// TwinCAT 3 PLC project TestRunner
// Title: TestRunner
// Company: Intecre Ltd
// ProjectVersion: 1.0.0.0
// Description: TcUnit test suites for the Intecre.File library. Not a library; activate it on a runtime (the usermode runtime works) to run the tests. The tests write their files to C:\TcUnit_IntecreFile.
// ProgramVersion: 3.1.4026.25
// libraries:
//   Tc2_Standard, * (Beckhoff Automation GmbH)
//   Tc2_System, * (Beckhoff Automation GmbH)
//   Tc2_Utilities, * (Beckhoff Automation GmbH)
//   TcUnit, * (www.tcunit.org)
//   Intecre.File, * (Intecre Ltd)
// project tree:
//   / MAIN.TcPOU, PlcTask.TcTTO
//   Helpers/ F_TestFilePath.TcPOU, ST_TestRecipe.TcDUT, T_TestDirectory.TcPOU, T_TestFile.TcPOU, TestFiles.TcGVL
//   Tests/ T_TxtFileWriter_Tests.TcPOU, T_CsvFileWriter_Tests.TcPOU, T_CsvFileReader_Tests.TcPOU, T_StructJsonFile_Tests.TcPOU, T_StructPersistence_Tests.TcPOU, T_CheckFileExists_Tests.TcPOU, ProjectInformation_Tests.TcPOU
// (motion and I/O tree: see PLC project intecre_file)
// real-time tasks:
//   TASK PlcTask: cycle T#10ms, priority 20, ADS port 350

CONFIGURATION TestRunner
    RESOURCE PLC ON TwinCAT3
        TASK PlcTask(INTERVAL := T#10ms, PRIORITY := 20);
        PROGRAM MAIN WITH PlcTask : MAIN;
    END_RESOURCE
END_CONFIGURATION

// ---- Helpers/ST_TestRecipe.TcDUT
TYPE ST_TestRecipe :
STRUCT
  Name : STRING(40);
  Speed : LREAL;
  Count : DINT;
  Enabled : BOOL;
END_STRUCT
END_TYPE

// ---- Helpers/TestFiles.TcGVL
{attribute 'qualified_only'}
VAR_GLOBAL CONSTANT
  DIRECTORY : T_MaxString := 'C:\TcUnit_IntecreFile';
  TIMEOUT : TIME := T#5S;
END_VAR

// ---- MAIN.TcPOU
PROGRAM MAIN
VAR
  testDirectory           : T_TestDirectory;
  suiteTxtFileWriter      : T_TxtFileWriter_Tests;
  suiteCsvFileWriter      : T_CsvFileWriter_Tests;
  suiteCsvFileReader      : T_CsvFileReader_Tests;
  suiteStructJsonFile     : T_StructJsonFile_Tests;
  suiteStructPersistence  : T_StructPersistence_Tests;
  suiteCheckFileExists    : T_CheckFileExists_Tests;
  suiteProjectInformation : ProjectInformation_Tests;
END_VAR

testDirectory();

IF NOT testDirectory.Ready THEN
  RETURN;
END_IF

TcUnit.RUN_IN_SEQUENCE();

END_PROGRAM

// ---- Helpers/T_TestDirectory.TcPOU
FUNCTION_BLOCK T_TestDirectory
VAR
  createDirectory : FB_CreateDir;
  requested : BOOL;
  _ready : BOOL;
END_VAR

IF _ready THEN
  RETURN;
END_IF

createDirectory(sNetId := '', sPathName := TestFiles.DIRECTORY, bExecute := TRUE);

IF requested AND NOT createDirectory.bBusy THEN
  _ready := TRUE;
END_IF

requested := TRUE;

PROPERTY Ready : BOOL
GET
Ready := _ready;
END_GET
END_PROPERTY

END_FUNCTION_BLOCK

// ---- Tests/T_TxtFileWriter_Tests.TcPOU
FUNCTION_BLOCK T_TxtFileWriter_Tests EXTENDS TcUnit.FB_TestSuite

Test_WriteLineEndsEachLineWithCrlf();
Test_WriteAddsToTheCurrentLine();
Test_AppendModeAddsToTheEndOfTheFile();
Test_OverwriteModeReplacesTheFile();
Test_ClearBufferDiscardsWhatWasWritten();
Test_ClearBufferReportsTheBufferIsClear();
Test_KeepsLinesLongerThan255Characters();
Test_MissingDirectoryGivesAnError();

METHOD PRIVATE Test_WriteLineEndsEachLineWithCrlf
VAR_INST
  writer : T_TxtFileWriter;
  testFile : T_TestFile;
  timeout : TON;
  step : INT;
END_VAR
IF NOT TcUnit.TEST_ORDERED(__POUNAME()) THEN
  RETURN;
END_IF

writer();
testFile();

timeout(IN := TRUE, PT := TestFiles.TIMEOUT);

IF timeout.Q THEN
  AssertTrue(Condition := FALSE, Message := 'the file operation did not finish in time');
  TEST_FINISHED_NAMED(__POUNAME());
  RETURN;
END_IF

CASE step OF

  0:

    writer.SetFileParams(FilePath := F_TestFilePath('txt_write_line.txt'));
    writer.WriteLine(Entry := 'first');
    writer.WriteLine(Entry := 'second');
    writer.WriteToFile();
    step := 10;

  10:

    IF writer.Busy THEN
      RETURN;
    END_IF

    AssertFalse(Condition := writer.Error, Message := 'file written without an error');
    testFile.Read(FilePath := F_TestFilePath('txt_write_line.txt'));
    step := 20;

  20:

    IF testFile.Busy THEN
      RETURN;
    END_IF

    AssertEquals_STRING(Expected := 'first$R$Nsecond$R$N', Actual := testFile.Text, Message := 'each line ends with CR LF');
    TEST_FINISHED_NAMED(__POUNAME());

END_CASE
END_METHOD

METHOD PRIVATE Test_WriteAddsToTheCurrentLine
VAR_INST
  writer : T_TxtFileWriter;
  testFile : T_TestFile;
  timeout : TON;
  step : INT;
END_VAR
IF NOT TcUnit.TEST_ORDERED(__POUNAME()) THEN
  RETURN;
END_IF

writer();
testFile();

timeout(IN := TRUE, PT := TestFiles.TIMEOUT);

IF timeout.Q THEN
  AssertTrue(Condition := FALSE, Message := 'the file operation did not finish in time');
  TEST_FINISHED_NAMED(__POUNAME());
  RETURN;
END_IF

CASE step OF

  0:

    writer.SetFileParams(FilePath := F_TestFilePath('txt_write.txt'));
    writer.Write(Entry := 'one');
    writer.Write(Entry := 'two');
    writer.NewLine();
    writer.WriteToFile();
    step := 10;

  10:

    IF writer.Busy THEN
      RETURN;
    END_IF

    AssertFalse(Condition := writer.Error, Message := 'file written without an error');
    testFile.Read(FilePath := F_TestFilePath('txt_write.txt'));
    step := 20;

  20:

    IF testFile.Busy THEN
      RETURN;
    END_IF

    AssertEquals_STRING(Expected := 'onetwo$R$N', Actual := testFile.Text, Message := 'Write adds to the line, NewLine ends it');
    TEST_FINISHED_NAMED(__POUNAME());

END_CASE
END_METHOD

METHOD PRIVATE Test_AppendModeAddsToTheEndOfTheFile
VAR_INST
  writer : T_TxtFileWriter;
  testFile : T_TestFile;
  timeout : TON;
  step : INT;
END_VAR
IF NOT TcUnit.TEST_ORDERED(__POUNAME()) THEN
  RETURN;
END_IF

writer();
testFile();

timeout(IN := TRUE, PT := TestFiles.TIMEOUT);

IF timeout.Q THEN
  AssertTrue(Condition := FALSE, Message := 'the file operation did not finish in time');
  TEST_FINISHED_NAMED(__POUNAME());
  RETURN;
END_IF

CASE step OF

  0:

    testFile.Write(FilePath := F_TestFilePath('txt_append.txt'), Content := 'existing$R$N');
    step := 5;

  5:

    IF testFile.Busy THEN
      RETURN;
    END_IF

    AssertFalse(Condition := testFile.Error, Message := 'existing file written');
    step := 6;

  6:

    writer.SetFileParams(FilePath := F_TestFilePath('txt_append.txt'));
    writer.SetFileOpenMode(Append := TRUE);
    writer.WriteLine(Entry := 'added');
    writer.WriteToFile();
    step := 10;

  10:

    IF writer.Busy THEN
      RETURN;
    END_IF

    AssertFalse(Condition := writer.Error, Message := 'file written without an error');
    testFile.Read(FilePath := F_TestFilePath('txt_append.txt'));
    step := 20;

  20:

    IF testFile.Busy THEN
      RETURN;
    END_IF

    AssertEquals_STRING(Expected := 'existing$R$Nadded$R$N', Actual := testFile.Text, Message := 'appended after the existing line');
    TEST_FINISHED_NAMED(__POUNAME());

END_CASE
END_METHOD

METHOD PRIVATE Test_OverwriteModeReplacesTheFile
VAR_INST
  writer : T_TxtFileWriter;
  testFile : T_TestFile;
  timeout : TON;
  step : INT;
END_VAR
IF NOT TcUnit.TEST_ORDERED(__POUNAME()) THEN
  RETURN;
END_IF

writer();
testFile();

timeout(IN := TRUE, PT := TestFiles.TIMEOUT);

IF timeout.Q THEN
  AssertTrue(Condition := FALSE, Message := 'the file operation did not finish in time');
  TEST_FINISHED_NAMED(__POUNAME());
  RETURN;
END_IF

CASE step OF

  0:

    testFile.Write(FilePath := F_TestFilePath('txt_overwrite.txt'), Content := 'old content$R$N');
    step := 5;

  5:

    IF testFile.Busy THEN
      RETURN;
    END_IF

    AssertFalse(Condition := testFile.Error, Message := 'existing file written');
    step := 6;

  6:

    writer.SetFileParams(FilePath := F_TestFilePath('txt_overwrite.txt'));
    writer.WriteLine(Entry := 'new');
    writer.WriteToFile();
    step := 10;

  10:

    IF writer.Busy THEN
      RETURN;
    END_IF

    AssertFalse(Condition := writer.Error, Message := 'file written without an error');
    testFile.Read(FilePath := F_TestFilePath('txt_overwrite.txt'));
    step := 20;

  20:

    IF testFile.Busy THEN
      RETURN;
    END_IF

    AssertEquals_STRING(Expected := 'new$R$N', Actual := testFile.Text, Message := 'the old content is gone');
    TEST_FINISHED_NAMED(__POUNAME());

END_CASE
END_METHOD

METHOD PRIVATE Test_ClearBufferDiscardsWhatWasWritten
VAR_INST
  writer : T_TxtFileWriter;
  testFile : T_TestFile;
  timeout : TON;
  step : INT;
END_VAR
IF NOT TcUnit.TEST_ORDERED(__POUNAME()) THEN
  RETURN;
END_IF

writer();
testFile();

timeout(IN := TRUE, PT := TestFiles.TIMEOUT);

IF timeout.Q THEN
  AssertTrue(Condition := FALSE, Message := 'the file operation did not finish in time');
  TEST_FINISHED_NAMED(__POUNAME());
  RETURN;
END_IF

CASE step OF

  0:

    writer.SetFileParams(FilePath := F_TestFilePath('txt_clear_buffer.txt'));
    writer.WriteLine(Entry := 'discarded');
    writer.ClearBuffer();
    writer.WriteLine(Entry := 'kept');
    writer.WriteToFile();
    step := 10;

  10:

    IF writer.Busy THEN
      RETURN;
    END_IF

    AssertFalse(Condition := writer.Error, Message := 'file written without an error');
    testFile.Read(FilePath := F_TestFilePath('txt_clear_buffer.txt'));
    step := 20;

  20:

    IF testFile.Busy THEN
      RETURN;
    END_IF

    AssertEquals_STRING(Expected := 'kept$R$N', Actual := testFile.Text, Message := 'only the line written after ClearBuffer');
    TEST_FINISHED_NAMED(__POUNAME());

END_CASE
END_METHOD

METHOD PRIVATE Test_ClearBufferReportsTheBufferIsClear
VAR_INST
  writer : T_TxtFileWriter;
END_VAR
IF NOT TcUnit.TEST_ORDERED(__POUNAME()) THEN
  RETURN;
END_IF

writer.WriteLine(Entry := 'line');
AssertTrue(Condition := writer.ClearBuffer(), Message := 'ClearBuffer returns TRUE');
AssertTrue(Condition := writer.BufferClear, Message := 'BufferClear after ClearBuffer');

TEST_FINISHED_NAMED(__POUNAME());
END_METHOD

METHOD PRIVATE Test_KeepsLinesLongerThan255Characters
VAR_INST
  writer : T_TxtFileWriter;
  testFile : T_TestFile;
  timeout : TON;
  step : INT;
  longLine : TxtFileString;
END_VAR
IF NOT TcUnit.TEST_ORDERED(__POUNAME()) THEN
  RETURN;
END_IF

writer();
testFile();

timeout(IN := TRUE, PT := TestFiles.TIMEOUT);

IF timeout.Q THEN
  AssertTrue(Condition := FALSE, Message := 'the file operation did not finish in time');
  TEST_FINISHED_NAMED(__POUNAME());
  RETURN;
END_IF

CASE step OF

  0:

    MEMSET(destAddr := ADR(longLine), fillByte := 16#41, n := 300);
    writer.SetFileParams(FilePath := F_TestFilePath('txt_long_line.txt'));
    writer.WriteLine(Entry := longLine);
    writer.WriteToFile();
    step := 10;

  10:

    IF writer.Busy THEN
      RETURN;
    END_IF

    testFile.Read(FilePath := F_TestFilePath('txt_long_line.txt'));
    step := 20;

  20:

    IF testFile.Busy THEN
      RETURN;
    END_IF

    AssertEquals_DINT(Expected := 302, Actual := testFile.Length, Message := '300 characters and CR LF');
    TEST_FINISHED_NAMED(__POUNAME());

END_CASE
END_METHOD

METHOD PRIVATE Test_MissingDirectoryGivesAnError
VAR_INST
  writer : T_TxtFileWriter;
  timeout : TON;
  step : INT;
END_VAR
IF NOT TcUnit.TEST_ORDERED(__POUNAME()) THEN
  RETURN;
END_IF

writer();

timeout(IN := TRUE, PT := TestFiles.TIMEOUT);

IF timeout.Q THEN
  AssertTrue(Condition := FALSE, Message := 'the file operation did not finish in time');
  TEST_FINISHED_NAMED(__POUNAME());
  RETURN;
END_IF

CASE step OF

  0:

    writer.SetFileParams(FilePath := F_TestFilePath('missing\file.txt'));
    writer.WriteLine(Entry := 'line');
    writer.WriteToFile();
    step := 10;

  10:

    IF writer.Busy THEN
      RETURN;
    END_IF

    AssertTrue(Condition := writer.Error, Message := 'a folder that does not exist gives an error');
    AssertTrue(Condition := writer.ErrorId <> 0, Message := 'with an error id');
    TEST_FINISHED_NAMED(__POUNAME());

END_CASE
END_METHOD

END_FUNCTION_BLOCK

// ---- Helpers/T_TestFile.TcPOU
FUNCTION_BLOCK T_TestFile
VAR
  fileOpen : FB_FileOpen;
  fileWrite : FB_FileWrite;
  fileRead : FB_FileRead;
  fileClose : FB_FileClose;
  fileDelete : FB_FileDelete;
  path : T_MaxString;
  textToWrite : STRING(2000);
  textRead : STRING(2000);
  startOfTextRead : T_MaxString;
  bytesRead : UDINT;
  request : (NoRequest, WriteRequest, ReadRequest, DeleteRequest);
  state : (Idle, Opening, Writing, Reading, Closing, Deleting);
  failed : BOOL;
END_VAR

CASE state OF

  Idle:

    IF request = DeleteRequest THEN
      state := Deleting;

    ELSIF request <> NoRequest THEN
      state := Opening;

    END_IF

  Opening:

    IF NOT fileOpen.bBusy AND fileOpen.bError THEN
      Finish(WithError := TRUE);

    ELSIF NOT fileOpen.bBusy AND (request = WriteRequest) THEN
      state := Writing;

    ELSIF NOT fileOpen.bBusy THEN
      state := Reading;

    END_IF

  Writing:

    IF NOT fileWrite.bBusy THEN
      failed := fileWrite.bError;
      state := Closing;
    END_IF

  Reading:

    IF NOT fileRead.bBusy THEN
      failed := fileRead.bError;
      bytesRead := fileRead.cbRead;
      MEMCPY(destAddr := ADR(startOfTextRead), srcAddr := ADR(textRead), n := SIZEOF(startOfTextRead) - 1);
      state := Closing;
    END_IF

  Closing:

    IF NOT fileClose.bBusy THEN
      Finish(WithError := failed OR fileClose.bError);
    END_IF

  Deleting:

    IF NOT fileDelete.bBusy THEN
      Finish(WithError := fileDelete.bError);
    END_IF

END_CASE

fileOpen(
  sNetId := '',
  sPathName := path,
  nMode := SEL(request = WriteRequest, FOPEN_MODEREAD OR FOPEN_MODEBINARY, FOPEN_MODEWRITE OR FOPEN_MODEBINARY),
  bExecute := state = Opening);

fileWrite(
  sNetId := '',
  hFile := fileOpen.hFile,
  pWriteBuff := ADR(textToWrite),
  cbWriteLen := TO_UDINT(LEN2(ADR(textToWrite))),
  bExecute := state = Writing);

fileRead(
  sNetId := '',
  hFile := fileOpen.hFile,
  pReadBuff := ADR(textRead),
  cbReadLen := SIZEOF(textRead) - 1,
  bExecute := state = Reading);

fileClose(
  sNetId := '',
  hFile := fileOpen.hFile,
  bExecute := state = Closing);

fileDelete(
  sNetId := '',
  sPathName := path,
  bExecute := state = Deleting);

PROPERTY Busy : BOOL
GET
Busy := request <> NoRequest;
END_GET
END_PROPERTY

METHOD Contains : BOOL
VAR_INPUT
  Part : T_MaxString;
END_VAR
VAR
  textLength : DINT;
  partLength : DINT;
  position : DINT;
END_VAR
textLength := TO_DINT(LEN2(ADR(textRead)));
partLength := TO_DINT(LEN2(ADR(Part)));

IF partLength = 0 THEN
  RETURN;
END_IF

FOR position := 0 TO textLength - partLength DO
  IF MEMCMP(pBuf1 := ADR(textRead) + TO_UDINT(position), pBuf2 := ADR(Part), n := TO_UDINT(partLength)) = 0 THEN
    Contains := TRUE;
    RETURN;
  END_IF
END_FOR
END_METHOD

METHOD Delete : BOOL
VAR_INPUT
  FilePath : T_MaxString;
END_VAR
IF Busy THEN
  RETURN;
END_IF

path := FilePath;
failed := FALSE;
request := DeleteRequest;
Delete := TRUE;
END_METHOD

PROPERTY Error : BOOL
GET
Error := failed AND NOT Busy;
END_GET
END_PROPERTY

METHOD PRIVATE Finish
VAR_INPUT
  WithError : BOOL;
END_VAR
failed := WithError;
request := NoRequest;
state := Idle;
END_METHOD

PROPERTY LastByte : BYTE // the last byte of the file the last Read read; 0 when it read nothing
GET // PUBLIC
IF bytesRead = 0 THEN
  RETURN;
END_IF

LastByte := textRead[bytesRead - 1];
END_GET
END_PROPERTY

PROPERTY Length : DINT
GET
Length := TO_DINT(LEN2(ADR(textRead)));
END_GET
END_PROPERTY

METHOD Read : BOOL
VAR_INPUT
  FilePath : T_MaxString;
END_VAR
IF Busy THEN
  RETURN;
END_IF

path := FilePath;
MEMSET(destAddr := ADR(textRead), fillByte := 0, n := SIZEOF(textRead));
MEMSET(destAddr := ADR(startOfTextRead), fillByte := 0, n := SIZEOF(startOfTextRead));
bytesRead := 0;
failed := FALSE;
request := ReadRequest;
Read := TRUE;
END_METHOD

PROPERTY Text : T_MaxString
GET
Text := startOfTextRead;
END_GET
END_PROPERTY

METHOD Write : BOOL
VAR_INPUT
  FilePath : T_MaxString;
  Content : STRING(2000);
END_VAR
IF Busy THEN
  RETURN;
END_IF

path := FilePath;
textToWrite := Content;
failed := FALSE;
request := WriteRequest;
Write := TRUE;
END_METHOD

END_FUNCTION_BLOCK

// ---- Helpers/F_TestFilePath.TcPOU
FUNCTION F_TestFilePath : T_MaxString
VAR_INPUT
  FileName : T_MaxString;
END_VAR

F_TestFilePath := CONCAT(CONCAT(TestFiles.DIRECTORY, '\'), FileName);

END_FUNCTION

// ---- Tests/T_CsvFileWriter_Tests.TcPOU
FUNCTION_BLOCK T_CsvFileWriter_Tests EXTENDS TcUnit.FB_TestSuite

Test_SeparatesFieldsWithCommas();
Test_SeparatesFieldsWithSemicolons();
Test_UnknownSeparatorFallsBackToSemicolon();
Test_AppendModeAddsRows();
Test_QuotesAFieldContainingTheSeparator();
Test_CountsRowsAndColumns();
Test_ClearBufferReportsTheBufferIsClear();

METHOD PRIVATE Test_SeparatesFieldsWithCommas
VAR_INST
  writer : T_CsvFileWriter;
  testFile : T_TestFile;
  timeout : TON;
  step : INT;
END_VAR
IF NOT TcUnit.TEST_ORDERED(__POUNAME()) THEN
  RETURN;
END_IF

writer();
testFile();

timeout(IN := TRUE, PT := TestFiles.TIMEOUT);

IF timeout.Q THEN
  AssertTrue(Condition := FALSE, Message := 'the file operation did not finish in time');
  TEST_FINISHED_NAMED(__POUNAME());
  RETURN;
END_IF

CASE step OF

  0:

    writer.SetFileParams(FilePath := F_TestFilePath('csv_commas.csv'), Separator := ASCI_COMMA);
    writer.AddStringField(sFieldString := 'a');
    writer.AddStringField(sFieldString := 'b');
    writer.NewLine();
    writer.AddStringField(sFieldString := 'c');
    writer.AddStringField(sFieldString := 'd');
    writer.WriteToFile();
    step := 10;

  10:

    IF writer.Busy THEN
      RETURN;
    END_IF

    AssertFalse(Condition := writer.Error, Message := 'file written without an error');
    testFile.Read(FilePath := F_TestFilePath('csv_commas.csv'));
    step := 20;

  20:

    IF testFile.Busy THEN
      RETURN;
    END_IF

    AssertEquals_STRING(Expected := 'a,b$R$Nc,d$R$N', Actual := testFile.Text, Message := 'two rows of two comma separated fields');
    TEST_FINISHED_NAMED(__POUNAME());

END_CASE
END_METHOD

METHOD PRIVATE Test_SeparatesFieldsWithSemicolons
VAR_INST
  writer : T_CsvFileWriter;
  testFile : T_TestFile;
  timeout : TON;
  step : INT;
END_VAR
IF NOT TcUnit.TEST_ORDERED(__POUNAME()) THEN
  RETURN;
END_IF

writer();
testFile();

timeout(IN := TRUE, PT := TestFiles.TIMEOUT);

IF timeout.Q THEN
  AssertTrue(Condition := FALSE, Message := 'the file operation did not finish in time');
  TEST_FINISHED_NAMED(__POUNAME());
  RETURN;
END_IF

CASE step OF

  0:

    writer.SetFileParams(FilePath := F_TestFilePath('csv_semicolons.csv'), Separator := ASCI_SEMI_COLON);
    writer.AddStringField(sFieldString := 'a');
    writer.AddStringField(sFieldString := 'b');
    writer.WriteToFile();
    step := 10;

  10:

    IF writer.Busy THEN
      RETURN;
    END_IF

    AssertFalse(Condition := writer.Error, Message := 'file written without an error');
    testFile.Read(FilePath := F_TestFilePath('csv_semicolons.csv'));
    step := 20;

  20:

    IF testFile.Busy THEN
      RETURN;
    END_IF

    AssertEquals_STRING(Expected := 'a;b$R$N', Actual := testFile.Text, Message := 'semicolon separated fields');
    TEST_FINISHED_NAMED(__POUNAME());

END_CASE
END_METHOD

METHOD PRIVATE Test_UnknownSeparatorFallsBackToSemicolon
VAR_INST
  writer : T_CsvFileWriter;
  testFile : T_TestFile;
  timeout : TON;
  step : INT;
END_VAR
IF NOT TcUnit.TEST_ORDERED(__POUNAME()) THEN
  RETURN;
END_IF

writer();
testFile();

timeout(IN := TRUE, PT := TestFiles.TIMEOUT);

IF timeout.Q THEN
  AssertTrue(Condition := FALSE, Message := 'the file operation did not finish in time');
  TEST_FINISHED_NAMED(__POUNAME());
  RETURN;
END_IF

CASE step OF

  0:

    writer.SetFileParams(FilePath := F_TestFilePath('csv_unknown_separator.csv'), Separator := 16#09);
    writer.AddStringField(sFieldString := 'a');
    writer.AddStringField(sFieldString := 'b');
    writer.WriteToFile();
    step := 10;

  10:

    IF writer.Busy THEN
      RETURN;
    END_IF

    AssertFalse(Condition := writer.Error, Message := 'file written without an error');
    testFile.Read(FilePath := F_TestFilePath('csv_unknown_separator.csv'));
    step := 20;

  20:

    IF testFile.Busy THEN
      RETURN;
    END_IF

    AssertEquals_STRING(Expected := 'a;b$R$N', Actual := testFile.Text, Message := 'a tab is not supported, so semicolon is used');
    TEST_FINISHED_NAMED(__POUNAME());

END_CASE
END_METHOD

METHOD PRIVATE Test_AppendModeAddsRows
VAR_INST
  writer : T_CsvFileWriter;
  testFile : T_TestFile;
  timeout : TON;
  step : INT;
END_VAR
IF NOT TcUnit.TEST_ORDERED(__POUNAME()) THEN
  RETURN;
END_IF

writer();
testFile();

timeout(IN := TRUE, PT := TestFiles.TIMEOUT);

IF timeout.Q THEN
  AssertTrue(Condition := FALSE, Message := 'the file operation did not finish in time');
  TEST_FINISHED_NAMED(__POUNAME());
  RETURN;
END_IF

CASE step OF

  0:

    testFile.Write(FilePath := F_TestFilePath('csv_append.csv'), Content := 'x,y$R$N');
    step := 5;

  5:

    IF testFile.Busy THEN
      RETURN;
    END_IF

    AssertFalse(Condition := testFile.Error, Message := 'existing file written');
    step := 6;

  6:

    writer.SetFileParams(FilePath := F_TestFilePath('csv_append.csv'), Separator := ASCI_COMMA);
    writer.SetFileOpenMode(Append := TRUE);
    writer.AddStringField(sFieldString := 'a');
    writer.AddStringField(sFieldString := 'b');
    writer.WriteToFile();
    step := 10;

  10:

    IF writer.Busy THEN
      RETURN;
    END_IF

    AssertFalse(Condition := writer.Error, Message := 'file written without an error');
    testFile.Read(FilePath := F_TestFilePath('csv_append.csv'));
    step := 20;

  20:

    IF testFile.Busy THEN
      RETURN;
    END_IF

    AssertEquals_STRING(Expected := 'x,y$R$Na,b$R$N', Actual := testFile.Text, Message := 'row appended after the existing row');
    TEST_FINISHED_NAMED(__POUNAME());

END_CASE
END_METHOD

METHOD PRIVATE Test_QuotesAFieldContainingTheSeparator
VAR_INST
  writer : T_CsvFileWriter;
  testFile : T_TestFile;
  timeout : TON;
  step : INT;
END_VAR
IF NOT TcUnit.TEST_ORDERED(__POUNAME()) THEN
  RETURN;
END_IF

writer();
testFile();

timeout(IN := TRUE, PT := TestFiles.TIMEOUT);

IF timeout.Q THEN
  AssertTrue(Condition := FALSE, Message := 'the file operation did not finish in time');
  TEST_FINISHED_NAMED(__POUNAME());
  RETURN;
END_IF

CASE step OF

  0:

    writer.SetFileParams(FilePath := F_TestFilePath('csv_quoted.csv'), Separator := ASCI_COMMA);
    writer.AddStringField(sFieldString := 'a,b');
    writer.AddStringField(sFieldString := 'c');
    writer.WriteToFile();
    step := 10;

  10:

    IF writer.Busy THEN
      RETURN;
    END_IF

    AssertFalse(Condition := writer.Error, Message := 'file written without an error');
    testFile.Read(FilePath := F_TestFilePath('csv_quoted.csv'));
    step := 20;

  20:

    IF testFile.Busy THEN
      RETURN;
    END_IF

    AssertEquals_STRING(Expected := '"a,b",c$R$N', Actual := testFile.Text, Message := 'a field holding the separator is quoted so the row keeps two fields');
    TEST_FINISHED_NAMED(__POUNAME());

END_CASE
END_METHOD

METHOD PRIVATE Test_CountsRowsAndColumns
VAR_INST
  writer : T_CsvFileWriter;
END_VAR
IF NOT TcUnit.TEST_ORDERED(__POUNAME()) THEN
  RETURN;
END_IF

writer.SetFileParams(FilePath := F_TestFilePath('csv_counts.csv'), Separator := ASCI_COMMA);
writer.AddStringField(sFieldString := 'a');
writer.AddStringField(sFieldString := 'b');
AssertEquals_UINT(Expected := 2, Actual := writer.Column, Message := 'two fields on the row');
AssertEquals_UINT(Expected := 0, Actual := writer.Row, Message := 'still on the first row');

writer.NewLine();
AssertEquals_UINT(Expected := 0, Actual := writer.Column, Message := 'column back to zero on a new line');
AssertEquals_UINT(Expected := 1, Actual := writer.Row, Message := 'second row');

TEST_FINISHED_NAMED(__POUNAME());
END_METHOD

METHOD PRIVATE Test_ClearBufferReportsTheBufferIsClear
VAR_INST
  writer : T_CsvFileWriter;
END_VAR
IF NOT TcUnit.TEST_ORDERED(__POUNAME()) THEN
  RETURN;
END_IF

writer.SetFileParams(FilePath := F_TestFilePath('csv_clear.csv'), Separator := ASCI_COMMA);
writer.AddStringField(sFieldString := 'a');
AssertTrue(Condition := writer.ClearBuffer(), Message := 'ClearBuffer returns TRUE');
AssertTrue(Condition := writer.BufferClear, Message := 'BufferClear after ClearBuffer');

TEST_FINISHED_NAMED(__POUNAME());
END_METHOD

END_FUNCTION_BLOCK

// ---- Tests/T_CsvFileReader_Tests.TcPOU
FUNCTION_BLOCK T_CsvFileReader_Tests EXTENDS TcUnit.FB_TestSuite

Test_ReadsEachFieldWithItsRowAndColumn();
Test_ReadsSemicolonSeparatedFields();
Test_KeepsFieldsLongerThan80Characters();
Test_MissingFileGivesAnError();

METHOD PRIVATE Test_KeepsFieldsLongerThan80Characters
VAR_INST
  reader : T_CsvFileReader;
  testFile : T_TestFile;
  timeout : TON;
  step : INT;
  content : STRING(2000);
  field : T_MaxString;
END_VAR
IF NOT TcUnit.TEST_ORDERED(__POUNAME()) THEN
  RETURN;
END_IF

reader();
testFile();

timeout(IN := TRUE, PT := TestFiles.TIMEOUT);

IF timeout.Q THEN
  AssertTrue(Condition := FALSE, Message := 'the file operation did not finish in time');
  TEST_FINISHED_NAMED(__POUNAME());
  RETURN;
END_IF

CASE step OF

  0:

    MEMSET(destAddr := ADR(content), fillByte := 16#41, n := 100);
    content[100] := 16#0D;
    content[101] := 16#0A;
    testFile.Write(FilePath := F_TestFilePath('csv_long_field.csv'), Content := content);
    step := 10;

  10:

    IF testFile.Busy THEN
      RETURN;
    END_IF

    AssertFalse(Condition := testFile.Error, Message := 'CSV file written for the test');
    reader.SetFileParams(FilePath := F_TestFilePath('csv_long_field.csv'), Separator := ASCI_COMMA);
    reader.GetFile();
    step := 20;

  20:

    IF reader.Busy THEN
      RETURN;
    END_IF

    AssertFalse(Condition := reader.Error, Message := 'file read without an error');
    AssertTrue(Condition := reader.ReadyForParsing, Message := 'ready for parsing');
    reader.NextField();
    field := reader.Field;
    AssertEquals_DINT(Expected := 100, Actual := TO_DINT(LEN2(ADR(field))), Message := 'all 100 characters of the field');
    TEST_FINISHED_NAMED(__POUNAME());

END_CASE
END_METHOD

METHOD PRIVATE Test_MissingFileGivesAnError
VAR_INST
  reader : T_CsvFileReader;
  testFile : T_TestFile;
  timeout : TON;
  step : INT;
END_VAR
IF NOT TcUnit.TEST_ORDERED(__POUNAME()) THEN
  RETURN;
END_IF

reader();
testFile();

timeout(IN := TRUE, PT := TestFiles.TIMEOUT);

IF timeout.Q THEN
  AssertTrue(Condition := FALSE, Message := 'the file operation did not finish in time');
  TEST_FINISHED_NAMED(__POUNAME());
  RETURN;
END_IF

CASE step OF

  0:

    testFile.Delete(FilePath := F_TestFilePath('csv_missing.csv'));
    step := 10;

  10:

    IF testFile.Busy THEN
      RETURN;
    END_IF

    reader.SetFileParams(FilePath := F_TestFilePath('csv_missing.csv'), Separator := ASCI_COMMA);
    reader.GetFile();
    step := 20;

  20:

    IF reader.Busy THEN
      RETURN;
    END_IF

    AssertTrue(Condition := reader.Error, Message := 'a missing file gives an error');
    AssertFalse(Condition := reader.FileExists, Message := 'FileExists is FALSE for a missing file');
    AssertFalse(Condition := reader.ReadyForParsing, Message := 'a missing file is not ready for parsing');
    TEST_FINISHED_NAMED(__POUNAME());

END_CASE
END_METHOD

METHOD PRIVATE Test_ReadsEachFieldWithItsRowAndColumn
VAR_INST
  reader : T_CsvFileReader;
  testFile : T_TestFile;
  timeout : TON;
  step : INT;
END_VAR
IF NOT TcUnit.TEST_ORDERED(__POUNAME()) THEN
  RETURN;
END_IF

reader();
testFile();

timeout(IN := TRUE, PT := TestFiles.TIMEOUT);

IF timeout.Q THEN
  AssertTrue(Condition := FALSE, Message := 'the file operation did not finish in time');
  TEST_FINISHED_NAMED(__POUNAME());
  RETURN;
END_IF

CASE step OF

  0:

    testFile.Write(FilePath := F_TestFilePath('csv_read.csv'), Content := 'a,b$R$Nc,d$R$N');
    step := 10;

  10:

    IF testFile.Busy THEN
      RETURN;
    END_IF

    AssertFalse(Condition := testFile.Error, Message := 'CSV file written for the test');
    reader.SetFileParams(FilePath := F_TestFilePath('csv_read.csv'), Separator := ASCI_COMMA);
    reader.GetFile();
    step := 20;

  20:

    IF reader.Busy THEN
      RETURN;
    END_IF

    AssertFalse(Condition := reader.Error, Message := 'file read without an error');
    AssertTrue(Condition := reader.ReadyForParsing, Message := 'ready for parsing');
    reader.NextField();
    AssertEquals_STRING(Expected := 'a', Actual := reader.Field, Message := 'field a');
    AssertEquals_UINT(Expected := 0, Actual := reader.Row, Message := 'row of a');
    AssertEquals_UINT(Expected := 0, Actual := reader.Column, Message := 'column of a');
    reader.NextField();
    AssertEquals_STRING(Expected := 'b', Actual := reader.Field, Message := 'field b');
    AssertEquals_UINT(Expected := 0, Actual := reader.Row, Message := 'row of b');
    AssertEquals_UINT(Expected := 1, Actual := reader.Column, Message := 'column of b');
    reader.NextField();
    AssertEquals_STRING(Expected := 'c', Actual := reader.Field, Message := 'field c');
    AssertEquals_UINT(Expected := 1, Actual := reader.Row, Message := 'row of c');
    AssertEquals_UINT(Expected := 0, Actual := reader.Column, Message := 'column of c');
    reader.NextField();
    AssertEquals_STRING(Expected := 'd', Actual := reader.Field, Message := 'field d');
    AssertEquals_UINT(Expected := 1, Actual := reader.Row, Message := 'row of d');
    AssertEquals_UINT(Expected := 1, Actual := reader.Column, Message := 'column of d');
    AssertFalse(Condition := reader.Eof, Message := 'not at the end on the last field');
    reader.NextField();
    AssertTrue(Condition := reader.Eof, Message := 'end of file after the last field');
    TEST_FINISHED_NAMED(__POUNAME());

END_CASE
END_METHOD

METHOD PRIVATE Test_ReadsSemicolonSeparatedFields
VAR_INST
  reader : T_CsvFileReader;
  testFile : T_TestFile;
  timeout : TON;
  step : INT;
END_VAR
IF NOT TcUnit.TEST_ORDERED(__POUNAME()) THEN
  RETURN;
END_IF

reader();
testFile();

timeout(IN := TRUE, PT := TestFiles.TIMEOUT);

IF timeout.Q THEN
  AssertTrue(Condition := FALSE, Message := 'the file operation did not finish in time');
  TEST_FINISHED_NAMED(__POUNAME());
  RETURN;
END_IF

CASE step OF

  0:

    testFile.Write(FilePath := F_TestFilePath('csv_read_semicolons.csv'), Content := 'a;b$R$N');
    step := 10;

  10:

    IF testFile.Busy THEN
      RETURN;
    END_IF

    AssertFalse(Condition := testFile.Error, Message := 'CSV file written for the test');
    reader.SetFileParams(FilePath := F_TestFilePath('csv_read_semicolons.csv'), Separator := ASCI_SEMI_COLON);
    reader.GetFile();
    step := 20;

  20:

    IF reader.Busy THEN
      RETURN;
    END_IF

    AssertFalse(Condition := reader.Error, Message := 'file read without an error');
    AssertTrue(Condition := reader.ReadyForParsing, Message := 'ready for parsing');
    reader.NextField();
    AssertEquals_STRING(Expected := 'a', Actual := reader.Field, Message := 'field a');
    AssertEquals_UINT(Expected := 0, Actual := reader.Row, Message := 'row of a');
    AssertEquals_UINT(Expected := 0, Actual := reader.Column, Message := 'column of a');
    reader.NextField();
    AssertEquals_STRING(Expected := 'b', Actual := reader.Field, Message := 'field b');
    AssertEquals_UINT(Expected := 0, Actual := reader.Row, Message := 'row of b');
    AssertEquals_UINT(Expected := 1, Actual := reader.Column, Message := 'column of b');
    TEST_FINISHED_NAMED(__POUNAME());

END_CASE
END_METHOD

END_FUNCTION_BLOCK

// ---- Tests/T_StructJsonFile_Tests.TcPOU
FUNCTION_BLOCK T_StructJsonFile_Tests EXTENDS TcUnit.FB_TestSuite

Test_WrittenStructReadsBackTheSame();
Test_ReadingAMissingFileGivesAnError();
Test_ReaderReadsAgainAfterAnErrorAndReset();
Test_ReaderRefusesAFileLongerThanJsonDocSize();
Test_WrittenFileEndsWithTheClosingBrace();

METHOD PRIVATE Test_ReaderReadsAgainAfterAnErrorAndReset
VAR_INST
  reader : T_StructFromJsonFileReader;
  testFile : T_TestFile;
  recipe : ST_TestRecipe;
  timeout : TON;
  step : INT;
END_VAR
IF NOT TcUnit.TEST_ORDERED(__POUNAME()) THEN
  RETURN;
END_IF

reader();
testFile();

timeout(IN := TRUE, PT := TestFiles.TIMEOUT);

IF timeout.Q THEN
  AssertTrue(Condition := FALSE, Message := 'the file operation did not finish in time');
  TEST_FINISHED_NAMED(__POUNAME());
  RETURN;
END_IF

CASE step OF

  0:

    testFile.Delete(FilePath := F_TestFilePath('json_after_reset.json'));
    step := 10;

  10:

    IF testFile.Busy THEN
      RETURN;
    END_IF

    reader.SetFileParams(
      FilePath := F_TestFilePath('json_after_reset.json'),
      StructureName := 'ST_TestRecipe',
      PointerToStructure := ADR(recipe),
      SizeOfStructure := SIZEOF(recipe));
    reader.ReadFromFile();
    step := 20;

  20:

    IF reader.Busy THEN
      RETURN;
    END_IF

    AssertTrue(Condition := reader.Error, Message := 'first read of a missing file fails');
    testFile.Write(FilePath := F_TestFilePath('json_after_reset.json'), Content := '{"Name":"from file","Speed":2.5,"Count":7,"Enabled":true}');
    step := 30;

  30:

    IF testFile.Busy THEN
      RETURN;
    END_IF

    reader.Reset();
    step := 40;

  40:

    reader.ReadFromFile();
    step := 50;

  50:

    IF reader.Busy THEN
      RETURN;
    END_IF

    AssertFalse(Condition := reader.Error, Message := 'the second read succeeds once the file exists');
    AssertEquals_DINT(Expected := 7, Actual := recipe.Count, Message := 'Count read from the file');
    TEST_FINISHED_NAMED(__POUNAME());

END_CASE
END_METHOD

METHOD PRIVATE Test_ReaderRefusesAFileLongerThanJsonDocSize
VAR_INST
  writer : T_TxtFileWriter;
  reader : T_StructFromJsonFileReader;
  testFile : T_TestFile;
  recipe : ST_TestRecipe;
  spaces : TxtFileString;
  spacesWritten : UDINT;
  timeout : TON;
  step : INT;
END_VAR
VAR CONSTANT
  SPACE : BYTE := 16#20;
  SPACES_PER_WRITE : UDINT := 200; // T_TxtFileWriter.Write keeps at most 255 characters a call
END_VAR
IF NOT TcUnit.TEST_ORDERED(__POUNAME()) THEN
  RETURN;
END_IF

writer();
reader();
testFile();

timeout(IN := TRUE, PT := TestFiles.TIMEOUT);

IF timeout.Q THEN
  AssertTrue(Condition := FALSE, Message := 'the file operation did not finish in time');
  TEST_FINISHED_NAMED(__POUNAME());
  RETURN;
END_IF

CASE step OF

  0:

    // arrange: JSON for the recipe, then spaces until the file is longer than JSON_DOC_SIZE
    MEMSET(destAddr := ADR(spaces), fillByte := SPACE, n := SPACES_PER_WRITE);
    writer.SetFileParams(FilePath := F_TestFilePath('json_too_long.json'));
    writer.Write(Entry := '{"Name":"from the long file","Speed":9.5,"Count":99,"Enabled":false}');

    WHILE spacesWritten <= Intecre_File.JsonParams.JSON_DOC_SIZE DO
      writer.Write(Entry := spaces);
      spacesWritten := spacesWritten + SPACES_PER_WRITE;
    END_WHILE

    writer.WriteToFile();
    step := 10;

  10:

    IF writer.Busy THEN
      RETURN;
    END_IF

    AssertFalse(Condition := writer.Error, Message := 'the long file was written');
    recipe.Name := 'unchanged';
    recipe.Speed := 1.5;
    recipe.Count := 1;
    recipe.Enabled := TRUE;
    reader.SetFileParams(
      FilePath := F_TestFilePath('json_too_long.json'),
      StructureName := 'ST_TestRecipe',
      PointerToStructure := ADR(recipe),
      SizeOfStructure := SIZEOF(recipe));

    // act
    reader.ReadFromFile();
    step := 20;

  20:

    IF reader.Busy THEN
      RETURN;
    END_IF

    // assert: the file is refused and the recipe is untouched
    AssertTrue(Condition := reader.Error, Message := 'a file longer than JSON_DOC_SIZE gives an error');
    AssertEquals_STRING(Expected := 'unchanged', Actual := recipe.Name, Message := 'Name untouched');
    AssertEquals_LREAL(Expected := 1.5, Actual := recipe.Speed, Delta := 0.0, Message := 'Speed untouched');
    AssertEquals_DINT(Expected := 1, Actual := recipe.Count, Message := 'Count untouched');
    AssertEquals_BOOL(Expected := TRUE, Actual := recipe.Enabled, Message := 'Enabled untouched');

    // the reader's settings are untouched if, after a Reset, it reads a short file into the same recipe
    testFile.Write(
      FilePath := F_TestFilePath('json_too_long.json'),
      Content := '{"Name":"from the short file","Speed":2.5,"Count":7,"Enabled":false}');
    step := 30;

  30:

    IF testFile.Busy THEN
      RETURN;
    END_IF

    AssertFalse(Condition := testFile.Error, Message := 'the short file was written');
    reader.Reset();
    step := 40;

  40:

    reader.ReadFromFile();
    step := 50;

  50:

    IF reader.Busy THEN
      RETURN;
    END_IF

    AssertFalse(Condition := reader.Error, Message := 'the reader reads a short file after the refusal and a Reset');
    AssertEquals_STRING(Expected := 'from the short file', Actual := recipe.Name, Message := 'structure name, address and size kept: Name read into the recipe');
    AssertEquals_DINT(Expected := 7, Actual := recipe.Count, Message := 'structure name, address and size kept: Count read into the recipe');
    TEST_FINISHED_NAMED(__POUNAME());

END_CASE
END_METHOD

METHOD PRIVATE Test_ReadingAMissingFileGivesAnError
VAR_INST
  reader : T_StructFromJsonFileReader;
  testFile : T_TestFile;
  recipe : ST_TestRecipe;
  timeout : TON;
  step : INT;
END_VAR
IF NOT TcUnit.TEST_ORDERED(__POUNAME()) THEN
  RETURN;
END_IF

reader();
testFile();

timeout(IN := TRUE, PT := TestFiles.TIMEOUT);

IF timeout.Q THEN
  AssertTrue(Condition := FALSE, Message := 'the file operation did not finish in time');
  TEST_FINISHED_NAMED(__POUNAME());
  RETURN;
END_IF

CASE step OF

  0:

    testFile.Delete(FilePath := F_TestFilePath('json_missing.json'));
    step := 10;

  10:

    IF testFile.Busy THEN
      RETURN;
    END_IF

    reader.SetFileParams(
      FilePath := F_TestFilePath('json_missing.json'),
      StructureName := 'ST_TestRecipe',
      PointerToStructure := ADR(recipe),
      SizeOfStructure := SIZEOF(recipe));
    reader.ReadFromFile();
    step := 20;

  20:

    IF reader.Busy THEN
      RETURN;
    END_IF

    AssertTrue(Condition := reader.Error, Message := 'a missing file gives an error');
    AssertFalse(Condition := reader.FileExists, Message := 'FileExists is FALSE');
    AssertFalse(Condition := reader.Done, Message := 'not done');
    TEST_FINISHED_NAMED(__POUNAME());

END_CASE
END_METHOD

METHOD PRIVATE Test_WrittenFileEndsWithTheClosingBrace
VAR_INST
  writer : T_StructToJsonFileWriter;
  testFile : T_TestFile;
  recipe : ST_TestRecipe;
  timeout : TON;
  step : INT;
END_VAR
VAR CONSTANT
  CLOSING_BRACE : BYTE := 16#7D; // }
END_VAR
IF NOT TcUnit.TEST_ORDERED(__POUNAME()) THEN
  RETURN;
END_IF

writer();
testFile();

timeout(IN := TRUE, PT := TestFiles.TIMEOUT);

IF timeout.Q THEN
  AssertTrue(Condition := FALSE, Message := 'the file operation did not finish in time');
  TEST_FINISHED_NAMED(__POUNAME());
  RETURN;
END_IF

CASE step OF

  0:

    // arrange
    recipe.Name := 'last byte';
    recipe.Speed := 3.25;
    recipe.Count := 5;
    recipe.Enabled := TRUE;
    writer.SetFileParams(
      FilePath := F_TestFilePath('json_last_byte.json'),
      StructureName := 'ST_TestRecipe',
      PointerToStructure := ADR(recipe),
      SizeOfStructure := SIZEOF(recipe));

    // act
    writer.WriteToFile();
    step := 10;

  10:

    IF writer.Busy THEN
      RETURN;
    END_IF

    AssertFalse(Condition := writer.Error, Message := 'struct written without an error');
    testFile.Read(FilePath := F_TestFilePath('json_last_byte.json'));
    step := 20;

  20:

    IF testFile.Busy THEN
      RETURN;
    END_IF

    // assert
    AssertFalse(Condition := testFile.Error, Message := 'the written file reads back');
    AssertEquals_BYTE(Expected := CLOSING_BRACE, Actual := testFile.LastByte, Message := 'the file ends with } and has no NUL after it');
    TEST_FINISHED_NAMED(__POUNAME());

END_CASE
END_METHOD

METHOD PRIVATE Test_WrittenStructReadsBackTheSame
VAR_INST
  writer : T_StructToJsonFileWriter;
  reader : T_StructFromJsonFileReader;
  original : ST_TestRecipe;
  copy : ST_TestRecipe;
  timeout : TON;
  step : INT;
END_VAR
IF NOT TcUnit.TEST_ORDERED(__POUNAME()) THEN
  RETURN;
END_IF

writer();
reader();

timeout(IN := TRUE, PT := TestFiles.TIMEOUT);

IF timeout.Q THEN
  AssertTrue(Condition := FALSE, Message := 'the file operation did not finish in time');
  TEST_FINISHED_NAMED(__POUNAME());
  RETURN;
END_IF

CASE step OF

  0:

    original.Name := 'recipe one';
    original.Speed := 12.5;
    original.Count := 42;
    original.Enabled := TRUE;
    writer.SetFileParams(
      FilePath := F_TestFilePath('json_round_trip.json'),
      StructureName := 'ST_TestRecipe',
      PointerToStructure := ADR(original),
      SizeOfStructure := SIZEOF(original));
    writer.WriteToFile();
    step := 10;

  10:

    IF writer.Busy THEN
      RETURN;
    END_IF

    AssertFalse(Condition := writer.Error, Message := 'struct written without an error');
    AssertTrue(Condition := writer.Done, Message := 'writer done');
    reader.SetFileParams(
      FilePath := F_TestFilePath('json_round_trip.json'),
      StructureName := 'ST_TestRecipe',
      PointerToStructure := ADR(copy),
      SizeOfStructure := SIZEOF(copy));
    reader.ReadFromFile();
    step := 20;

  20:

    IF reader.Busy THEN
      RETURN;
    END_IF

    AssertFalse(Condition := reader.Error, Message := 'struct read without an error');
    AssertTrue(Condition := reader.Done, Message := 'reader done');
    AssertEquals_STRING(Expected := original.Name, Actual := copy.Name, Message := 'Name');
    AssertEquals_LREAL(Expected := original.Speed, Actual := copy.Speed, Delta := 1.0E-9, Message := 'Speed');
    AssertEquals_DINT(Expected := original.Count, Actual := copy.Count, Message := 'Count');
    AssertEquals_BOOL(Expected := original.Enabled, Actual := copy.Enabled, Message := 'Enabled');
    TEST_FINISHED_NAMED(__POUNAME());

END_CASE
END_METHOD

END_FUNCTION_BLOCK

// ---- Tests/T_StructPersistence_Tests.TcPOU
FUNCTION_BLOCK T_StructPersistence_Tests EXTENDS TcUnit.FB_TestSuite

Test_CreatesTheFileWhenItDoesNotExist();
Test_ReadsAnExistingFileIntoTheStruct();
Test_ReadsAgainAfterAFailedRead();
Test_WriteToFileSavesTheCurrentStruct();
Test_AutoWritesAfterTheStructChanges();
Test_CreatesAFileWithAPathLongerThan80Characters();

METHOD PRIVATE Test_CreatesTheFileWhenItDoesNotExist
VAR_INST
  persistence : T_StructPersistence;
  options : ST_PersistenceOptions;
  recipe : ST_TestRecipe;
  testFile : T_TestFile;
  timeout : TON;
  settle : TON;
  step : INT;
END_VAR
IF NOT TcUnit.TEST_ORDERED(__POUNAME()) THEN
  RETURN;
END_IF

testFile();

IF step >= 20 THEN
  persistence(Options := options);
END_IF

timeout(IN := TRUE, PT := TestFiles.TIMEOUT);

IF timeout.Q THEN
  AssertTrue(Condition := FALSE, Message := 'the file operation did not finish in time');
  TEST_FINISHED_NAMED(__POUNAME());
  RETURN;
END_IF

CASE step OF

  0:

    testFile.Delete(FilePath := F_TestFilePath('persist_create.json'));
    step := 10;

  10:

    IF testFile.Busy THEN
      RETURN;
    END_IF

    recipe.Count := 5;
    options.AddressOfStruct := ADR(recipe);
    options.SizeOfStruct := SIZEOF(recipe);
    options.NameOfStructureType := 'ST_TestRecipe';
    options.FilePath := F_TestFilePath('persist_create.json');
    options.CreateFileIfDoesntExist := TRUE;
    options.AutoWriteOnDifference := FALSE;
    options.AutoWriteCheckTime := T#200MS;
    options.AutoWriteDebounceTime := T#200MS;
    step := 20;

  20:

    IF NOT persistence.FileCreated THEN
      RETURN;
    END_IF

    AssertTrue(Condition := persistence.WriteSuccess, Message := 'write reported');
    testFile.Read(FilePath := F_TestFilePath('persist_create.json'));
    step := 30;

  30:

    IF testFile.Busy THEN
      RETURN;
    END_IF

    AssertTrue(Condition := testFile.Contains('"Count":5'), Message := 'the new file holds the struct');
    TEST_FINISHED_NAMED(__POUNAME());

END_CASE
END_METHOD

METHOD PRIVATE Test_ReadsAnExistingFileIntoTheStruct
VAR_INST
  persistence : T_StructPersistence;
  options : ST_PersistenceOptions;
  recipe : ST_TestRecipe;
  testFile : T_TestFile;
  timeout : TON;
  settle : TON;
  step : INT;
END_VAR
IF NOT TcUnit.TEST_ORDERED(__POUNAME()) THEN
  RETURN;
END_IF

testFile();

IF step >= 20 THEN
  persistence(Options := options);
END_IF

timeout(IN := TRUE, PT := TestFiles.TIMEOUT);

IF timeout.Q THEN
  AssertTrue(Condition := FALSE, Message := 'the file operation did not finish in time');
  TEST_FINISHED_NAMED(__POUNAME());
  RETURN;
END_IF

CASE step OF

  0:

    testFile.Write(FilePath := F_TestFilePath('persist_read.json'), Content := '{"Name":"from file","Speed":2.5,"Count":7,"Enabled":true}');
    step := 10;

  10:

    IF testFile.Busy THEN
      RETURN;
    END_IF

    options.AddressOfStruct := ADR(recipe);
    options.SizeOfStruct := SIZEOF(recipe);
    options.NameOfStructureType := 'ST_TestRecipe';
    options.FilePath := F_TestFilePath('persist_read.json');
    options.CreateFileIfDoesntExist := TRUE;
    options.AutoWriteOnDifference := FALSE;
    options.AutoWriteCheckTime := T#200MS;
    options.AutoWriteDebounceTime := T#200MS;
    step := 20;

  20:

    IF NOT persistence.ReadSuccess THEN
      RETURN;
    END_IF

    AssertEquals_STRING(Expected := 'from file', Actual := recipe.Name, Message := 'Name read from the file');
    AssertEquals_DINT(Expected := 7, Actual := recipe.Count, Message := 'Count read from the file');
    AssertFalse(Condition := persistence.FileCreated, Message := 'an existing file is not created again');
    TEST_FINISHED_NAMED(__POUNAME());

END_CASE
END_METHOD

METHOD PRIVATE Test_ReadsAgainAfterAFailedRead
VAR_INST
  persistence : T_StructPersistence;
  options : ST_PersistenceOptions;
  recipe : ST_TestRecipe;
  testFile : T_TestFile;
  timeout : TON;
  settle : TON;
  step : INT;
END_VAR
IF NOT TcUnit.TEST_ORDERED(__POUNAME()) THEN
  RETURN;
END_IF

testFile();

IF step >= 20 THEN
  persistence(Options := options);
END_IF

timeout(IN := TRUE, PT := TestFiles.TIMEOUT);

IF timeout.Q THEN
  AssertTrue(Condition := FALSE, Message := 'the file operation did not finish in time');
  TEST_FINISHED_NAMED(__POUNAME());
  RETURN;
END_IF

CASE step OF

  0:

    testFile.Delete(FilePath := F_TestFilePath('persist_read_again.json'));
    step := 10;

  10:

    IF testFile.Busy THEN
      RETURN;
    END_IF

    options.AddressOfStruct := ADR(recipe);
    options.SizeOfStruct := SIZEOF(recipe);
    options.NameOfStructureType := 'ST_TestRecipe';
    options.FilePath := F_TestFilePath('persist_read_again.json');
    options.CreateFileIfDoesntExist := FALSE;
    options.AutoWriteOnDifference := FALSE;
    options.AutoWriteCheckTime := T#200MS;
    options.AutoWriteDebounceTime := T#200MS;
    step := 20;

  20:

    settle(IN := TRUE, PT := T#500MS);

    IF NOT settle.Q THEN
      RETURN;
    END_IF

    AssertFalse(Condition := persistence.ReadSuccess, Message := 'the first read fails while the file is missing');
    testFile.Write(FilePath := F_TestFilePath('persist_read_again.json'), Content := '{"Name":"from file","Speed":2.5,"Count":7,"Enabled":true}');
    step := 30;

  30:

    IF testFile.Busy THEN
      RETURN;
    END_IF

    AssertTrue(Condition := persistence.ReadFromFile(), Message := 'read requested');
    step := 40;

  40:

    IF NOT persistence.ReadSuccess THEN
      RETURN;
    END_IF

    AssertEquals_DINT(Expected := 7, Actual := recipe.Count, Message := 'Count read from the file');
    TEST_FINISHED_NAMED(__POUNAME());

END_CASE
END_METHOD

METHOD PRIVATE Test_WriteToFileSavesTheCurrentStruct
VAR_INST
  persistence : T_StructPersistence;
  options : ST_PersistenceOptions;
  recipe : ST_TestRecipe;
  testFile : T_TestFile;
  timeout : TON;
  settle : TON;
  step : INT;
END_VAR
IF NOT TcUnit.TEST_ORDERED(__POUNAME()) THEN
  RETURN;
END_IF

testFile();

IF step >= 20 THEN
  persistence(Options := options);
END_IF

timeout(IN := TRUE, PT := TestFiles.TIMEOUT);

IF timeout.Q THEN
  AssertTrue(Condition := FALSE, Message := 'the file operation did not finish in time');
  TEST_FINISHED_NAMED(__POUNAME());
  RETURN;
END_IF

CASE step OF

  0:

    testFile.Write(FilePath := F_TestFilePath('persist_write.json'), Content := '{"Name":"from file","Speed":2.5,"Count":7,"Enabled":true}');
    step := 10;

  10:

    IF testFile.Busy THEN
      RETURN;
    END_IF

    options.AddressOfStruct := ADR(recipe);
    options.SizeOfStruct := SIZEOF(recipe);
    options.NameOfStructureType := 'ST_TestRecipe';
    options.FilePath := F_TestFilePath('persist_write.json');
    options.CreateFileIfDoesntExist := TRUE;
    options.AutoWriteOnDifference := FALSE;
    options.AutoWriteCheckTime := T#200MS;
    options.AutoWriteDebounceTime := T#200MS;
    step := 20;

  20:

    IF NOT persistence.ReadSuccess THEN
      RETURN;
    END_IF

    recipe.Count := 21;
    AssertTrue(Condition := persistence.WriteToFile(), Message := 'write requested');
    step := 30;

  30:

    IF NOT persistence.WriteSuccess THEN
      RETURN;
    END_IF

    testFile.Read(FilePath := F_TestFilePath('persist_write.json'));
    step := 40;

  40:

    IF testFile.Busy THEN
      RETURN;
    END_IF

    AssertTrue(Condition := testFile.Contains('"Count":21'), Message := 'the file holds the changed struct');
    TEST_FINISHED_NAMED(__POUNAME());

END_CASE
END_METHOD

METHOD PRIVATE Test_AutoWritesAfterTheStructChanges
VAR_INST
  persistence : T_StructPersistence;
  options : ST_PersistenceOptions;
  recipe : ST_TestRecipe;
  testFile : T_TestFile;
  timeout : TON;
  settle : TON;
  step : INT;
END_VAR
IF NOT TcUnit.TEST_ORDERED(__POUNAME()) THEN
  RETURN;
END_IF

testFile();

IF step >= 20 THEN
  persistence(Options := options);
END_IF

timeout(IN := TRUE, PT := TestFiles.TIMEOUT);

IF timeout.Q THEN
  AssertTrue(Condition := FALSE, Message := 'the file operation did not finish in time');
  TEST_FINISHED_NAMED(__POUNAME());
  RETURN;
END_IF

CASE step OF

  0:

    testFile.Write(FilePath := F_TestFilePath('persist_auto_write.json'), Content := '{"Name":"from file","Speed":2.5,"Count":7,"Enabled":true}');
    step := 10;

  10:

    IF testFile.Busy THEN
      RETURN;
    END_IF

    options.AddressOfStruct := ADR(recipe);
    options.SizeOfStruct := SIZEOF(recipe);
    options.NameOfStructureType := 'ST_TestRecipe';
    options.FilePath := F_TestFilePath('persist_auto_write.json');
    options.CreateFileIfDoesntExist := TRUE;
    options.AutoWriteOnDifference := TRUE;
    options.AutoWriteCheckTime := T#200MS;
    options.AutoWriteDebounceTime := T#200MS;
    step := 20;

  20:

    IF NOT persistence.ReadSuccess THEN
      RETURN;
    END_IF

    recipe.Count := 33;
    step := 30;

  30:

    settle(IN := TRUE, PT := T#1500MS);

    IF NOT settle.Q THEN
      RETURN;
    END_IF

    testFile.Read(FilePath := F_TestFilePath('persist_auto_write.json'));
    step := 40;

  40:

    IF testFile.Busy THEN
      RETURN;
    END_IF

    AssertTrue(Condition := testFile.Contains('"Count":33'), Message := 'the change was written without a WriteToFile call');
    TEST_FINISHED_NAMED(__POUNAME());

END_CASE
END_METHOD

METHOD PRIVATE Test_CreatesAFileWithAPathLongerThan80Characters
VAR_INST
  persistence : T_StructPersistence;
  options : ST_PersistenceOptions;
  recipe : ST_TestRecipe;
  testFile : T_TestFile;
  timeout : TON;
  settle : TON;
  step : INT;
END_VAR
IF NOT TcUnit.TEST_ORDERED(__POUNAME()) THEN
  RETURN;
END_IF

testFile();

IF step >= 20 THEN
  persistence(Options := options);
END_IF

timeout(IN := TRUE, PT := TestFiles.TIMEOUT);

IF timeout.Q THEN
  AssertTrue(Condition := FALSE, Message := 'the file operation did not finish in time');
  TEST_FINISHED_NAMED(__POUNAME());
  RETURN;
END_IF

CASE step OF

  0:

    testFile.Delete(FilePath := F_TestFilePath('a_file_name_that_makes_the_whole_path_longer_than_eighty_characters.json'));
    step := 10;

  10:

    IF testFile.Busy THEN
      RETURN;
    END_IF

    recipe.Count := 8;
    options.AddressOfStruct := ADR(recipe);
    options.SizeOfStruct := SIZEOF(recipe);
    options.NameOfStructureType := 'ST_TestRecipe';
    options.FilePath := F_TestFilePath('a_file_name_that_makes_the_whole_path_longer_than_eighty_characters.json');
    options.CreateFileIfDoesntExist := TRUE;
    options.AutoWriteOnDifference := FALSE;
    options.AutoWriteCheckTime := T#200MS;
    options.AutoWriteDebounceTime := T#200MS;
    step := 20;

  20:

    IF NOT persistence.WriteSuccess THEN
      RETURN;
    END_IF

    testFile.Read(FilePath := F_TestFilePath('a_file_name_that_makes_the_whole_path_longer_than_eighty_characters.json'));
    step := 30;

  30:

    IF testFile.Busy THEN
      RETURN;
    END_IF

    AssertFalse(Condition := testFile.Error, Message := 'the file is at the full path');
    AssertTrue(Condition := testFile.Contains('"Count":8'), Message := 'and holds the struct');
    TEST_FINISHED_NAMED(__POUNAME());

END_CASE
END_METHOD

END_FUNCTION_BLOCK

// ---- Tests/T_CheckFileExists_Tests.TcPOU
FUNCTION_BLOCK T_CheckFileExists_Tests EXTENDS TcUnit.FB_TestSuite

Test_FindsAnExistingFile();
Test_ReportsAMissingFile();
Test_FindsAFileWithAPathLongerThan80Characters();

METHOD PRIVATE Test_FindsAnExistingFile
VAR_INST
  checker : T_CheckFileExists;
  testFile : T_TestFile;
  timeout : TON;
  step : INT;
END_VAR
IF NOT TcUnit.TEST_ORDERED(__POUNAME()) THEN
  RETURN;
END_IF

checker();
testFile();

timeout(IN := TRUE, PT := TestFiles.TIMEOUT);

IF timeout.Q THEN
  AssertTrue(Condition := FALSE, Message := 'the file operation did not finish in time');
  TEST_FINISHED_NAMED(__POUNAME());
  RETURN;
END_IF

CASE step OF

  0:

    testFile.Write(FilePath := F_TestFilePath('exists.txt'), Content := 'x');
    step := 10;

  10:

    IF testFile.Busy THEN
      RETURN;
    END_IF

    checker.Check(Path := F_TestFilePath('exists.txt'));
    step := 20;

  20:

    IF checker.Busy THEN
      RETURN;
    END_IF

    AssertEquals_BOOL(Expected := TRUE, Actual := checker.FileExists, Message := 'an existing file is found');
    TEST_FINISHED_NAMED(__POUNAME());

END_CASE
END_METHOD

METHOD PRIVATE Test_ReportsAMissingFile
VAR_INST
  checker : T_CheckFileExists;
  testFile : T_TestFile;
  timeout : TON;
  step : INT;
END_VAR
IF NOT TcUnit.TEST_ORDERED(__POUNAME()) THEN
  RETURN;
END_IF

checker();
testFile();

timeout(IN := TRUE, PT := TestFiles.TIMEOUT);

IF timeout.Q THEN
  AssertTrue(Condition := FALSE, Message := 'the file operation did not finish in time');
  TEST_FINISHED_NAMED(__POUNAME());
  RETURN;
END_IF

CASE step OF

  0:

    testFile.Delete(FilePath := F_TestFilePath('does_not_exist.txt'));
    step := 10;

  10:

    IF testFile.Busy THEN
      RETURN;
    END_IF

    checker.Check(Path := F_TestFilePath('does_not_exist.txt'));
    step := 20;

  20:

    IF checker.Busy THEN
      RETURN;
    END_IF

    AssertEquals_BOOL(Expected := FALSE, Actual := checker.FileExists, Message := 'a missing file is not found');
    TEST_FINISHED_NAMED(__POUNAME());

END_CASE
END_METHOD

METHOD PRIVATE Test_FindsAFileWithAPathLongerThan80Characters
VAR_INST
  checker : T_CheckFileExists;
  testFile : T_TestFile;
  timeout : TON;
  step : INT;
END_VAR
IF NOT TcUnit.TEST_ORDERED(__POUNAME()) THEN
  RETURN;
END_IF

checker();
testFile();

timeout(IN := TRUE, PT := TestFiles.TIMEOUT);

IF timeout.Q THEN
  AssertTrue(Condition := FALSE, Message := 'the file operation did not finish in time');
  TEST_FINISHED_NAMED(__POUNAME());
  RETURN;
END_IF

CASE step OF

  0:

    testFile.Write(FilePath := F_TestFilePath('a_file_name_that_makes_the_whole_path_longer_than_eighty_characters.json.txt'), Content := 'x');
    step := 10;

  10:

    IF testFile.Busy THEN
      RETURN;
    END_IF

    checker.Check(Path := F_TestFilePath('a_file_name_that_makes_the_whole_path_longer_than_eighty_characters.json.txt'));
    step := 20;

  20:

    IF checker.Busy THEN
      RETURN;
    END_IF

    AssertEquals_BOOL(Expected := TRUE, Actual := checker.FileExists, Message := 'a path longer than 80 characters is checked in full');
    TEST_FINISHED_NAMED(__POUNAME());

END_CASE
END_METHOD

END_FUNCTION_BLOCK

// ---- Tests/ProjectInformation_Tests.TcPOU
FUNCTION_BLOCK ProjectInformation_Tests EXTENDS TcUnit.FB_TestSuite

Test_TitleAndCompany();
Test_VersionIsOnePointThree();

METHOD PRIVATE Test_TitleAndCompany
TcUnit.TEST(__POUNAME());

AssertEquals_WSTRING(Expected := "Intecre.File", Actual := Intecre_File.F_GetTitle(), Message := 'library title');
AssertEquals_WSTRING(Expected := "Intecre Ltd", Actual := Intecre_File.F_GetCompany(), Message := 'library company');

TEST_FINISHED_NAMED(__POUNAME());
END_METHOD

METHOD PRIVATE Test_VersionIsOnePointThree
VAR
  version : ST_LibVersion;
END_VAR
TcUnit.TEST(__POUNAME());

version := Intecre_File.F_GetVersion();
AssertEquals_STRING(Expected := '1.3.1.0', Actual := version.sVersion, Message := 'library version string');
AssertEquals_UINT(Expected := 1, Actual := version.iMajor, Message := 'major version');
AssertEquals_UINT(Expected := 3, Actual := version.iMinor, Message := 'minor version');

TEST_FINISHED_NAMED(__POUNAME());
END_METHOD

END_FUNCTION_BLOCK
